(* IEC 61131-3 sources: sis-interlock-demo/tests/POUs/Generated/FB_CemGen03_Test, 3 files *)

(* ---- FB_CemGen03_Test.decl.st ---- *)
// AUTO-GENERATED by cemgen 1.0.0 — не редактировать: правьте матрицу и запустите
//   python -m cemgen generate <файл матрицы .csv или .xlsx>
// Матрица: SIS-V101-CEM, объект V-101, ревизия B от 2026-10-19, SHA-256 сетки df2ed4841a9453ca
// Назначение: набор coUnit: сценарии по матрице SIS-V101-CEM, тесты 81–83 (DESIGN.md, 12.4).
//             Ожидаемые значения — эталонная модель cemgen. Стенд FB_SisHarness — по экземпляру на
//             тест.
// Автор:      kr0nsch; код — генератор cemgen
// Версия:     1.0.0
// Документ:   docs/DESIGN.md, раздел «10. Генератор cemgen»; docs/cause_effect_matrix.md
// ВНИМАНИЕ:   код демонстрационный и не предназначен для систем безопасности. Реальная ПАЗ требует
//             определения SIL, сертифицированных аппаратных и программных средств и валидации по
//             ГОСТ Р МЭК 61511.
FUNCTION_BLOCK FB_CemGen03_Test EXTENDS coUnit.FB_TestSuite
VAR
    fbH001 : FB_SisHarness;   // Matrix_Start_TrippedUntilReset
    fbH002 : FB_SisHarness;   // Matrix_FirstOutSimultaneous_LowestIndex
    fbH003 : FB_SisHarness;   // Matrix_GeneratedCfg_PassesChecks
END_VAR

(* ---- FirstOutSimultaneousLowestIndex.method.decl.st ---- *)
// AUTO-GENERATED by cemgen 1.0.0 — не редактировать: правьте матрицу и запустите
//   python -m cemgen generate <файл матрицы .csv или .xlsx>
// Матрица: SIS-V101-CEM, объект V-101, ревизия B от 2026-10-19, SHA-256 сетки df2ed4841a9453ca
// Назначение: тест Matrix_FirstOutSimultaneous_LowestIndex набора FB_CemGen03_Test (сценарий по
//             матрице, DESIGN.md, 12.4).
// Автор:      kr0nsch; код — генератор cemgen
// Версия:     1.0.0
// Документ:   docs/DESIGN.md, раздел «10. Генератор cemgen»; docs/cause_effect_matrix.md
// ВНИМАНИЕ:   код демонстрационный и не предназначен для систем безопасности. Реальная ПАЗ требует
//             определения SIL, сертифицированных аппаратных и программных средств и валидации по
//             ГОСТ Р МЭК 61511.
// Одновременная фиксация PSHH101 и LSHH102 (без общих каналов) в одном вызове: требования подаются со
// сдвигом на разницу задержек → первопричина — младшая причина, в маске первопричины обе.
METHOD PRIVATE FirstOutSimultaneousLowestIndex
VAR
    xArmed : BOOL;   // стенд взведён: все следствия под напряжением после сброса
END_VAR

(* ---- GeneratedCfgPassesChecks.method.decl.st ---- *)
// AUTO-GENERATED by cemgen 1.0.0 — не редактировать: правьте матрицу и запустите
//   python -m cemgen generate <файл матрицы .csv или .xlsx>
// Матрица: SIS-V101-CEM, объект V-101, ревизия B от 2026-10-19, SHA-256 сетки df2ed4841a9453ca
// Назначение: тест Matrix_GeneratedCfg_PassesChecks набора FB_CemGen03_Test (сценарий по матрице,
//             DESIGN.md, 12.4).
// Автор:      kr0nsch; код — генератор cemgen
// Версия:     1.0.0
// Документ:   docs/DESIGN.md, раздел «10. Генератор cemgen»; docs/cause_effect_matrix.md
// ВНИМАНИЕ:   код демонстрационный и не предназначен для систем безопасности. Реальная ПАЗ требует
//             определения SIL, сертифицированных аппаратных и программных средств и валидации по
//             ГОСТ Р МЭК 61511.
// Сгенерированная конфигурация: F_CemCrc(CEM_CFG) = 16#CD40 = CEM_CFG.wMatrixCrc, F_CemCheckCfg без
// ошибок; после взвода нет ошибок конфигурации у матрицы и у групп голосования.
METHOD PRIVATE GeneratedCfgPassesChecks
VAR
    stCfg  : ST_CemCfg;      // копия GVL_SisCfg.CEM_CFG
    wCrc   : WORD;           // CRC сгенерированной матрицы
    wErr   : WORD;           // биты ошибок конфигурации матрицы
    xArmed : BOOL;           // стенд взведён: все следствия под напряжением после сброса
    stVs   : ST_VotingSts;   // копия состояния группы голосования
END_VAR
